(* IEC 61131-3 sources: plc-process-lib/tools/demo/src/POUs/FB_DemoLevelLoop, 2 files *)

(* ---- FB_DemoLevelLoop.decl.st ---- *)
// Назначение: сценарий A демонстрационного прогона — контур уровня по примеру 17.3 контракта:
//             LT (PL.FB_AnalogInput, 4–20 мА, 0..5 м) -> LIC (PL.FB_PID, Direct, обратный расчёт
//             по фактическому заданию ПЧ) -> насос с ПЧ (PL.FB_MotorVfd, мин. 20 %). Объект —
//             модель ёмкости на ST: баланс объёма, подача насоса пропорциональна скорости, ПЧ
//             разгоняется с рампой. Сценарий: 5 с — пуск насоса (слежение ПИД снимается без
//             рывка); 40 с — задание 2,5 -> 1,5 м (выход упирается в 100 %, интегратор не
//             накапливается); 95 с — приток 120 -> 210 м3/ч. Ёмкость и параметры вымышленные.
//             Коды событий: 1 — пуск насоса, 2 — ступень задания, 3 — ступень притока.
// Автор:      kr0nsch
// Версия:     0.1.0
// Документ:   docs/API.md, пример 17.3; tools/demo/README.md
FUNCTION_BLOCK FB_DemoLevelLoop
VAR_INPUT
    lrT_s  : LREAL;   // время от старта сценария, с
    lrDt_s : LREAL;   // шаг времени этого цикла, с
END_VAR
VAR_OUTPUT
    xDone : BOOL;     // сценарий завершён, журнал записан
END_VAR
VAR CONSTANT
    LEVEL_SPAN_M   : REAL := 5.0;       // шкала датчика: 4 мА = 0 м, 20 мА = 5 м
    MA_LO          : REAL := 4.0;       // ток начала шкалы, мА
    MA_SPAN        : REAL := 16.0;      // диапазон тока шкалы, мА
    AREA_M2        : LREAL := 1.5;      // площадь сечения ёмкости, м2
    LEVEL0_M       : LREAL := 2.3;      // начальный уровень, м
    Q_PUMP_MAX_M3H : REAL := 300.0;     // подача насоса при 100 % скорости, м3/ч (линейная модель)
    Q_IN_BASE_M3H  : REAL := 120.0;     // приток до возмущения, м3/ч
    Q_IN_SURGE_M3H : REAL := 210.0;     // приток после возмущения, м3/ч
    VFD_RAMP_PCTPS : REAL := 25.0;      // рампа ПЧ (модель привода), %/с
    S_PER_H        : LREAL := 3600.0;   // секунд в часе
    PCT_FULL       : REAL := 100.0;     // 100 %
    SP0_M          : REAL := 2.5;       // задание до ступени, м
    SP1_M          : REAL := 1.5;       // задание после ступени, м
    T_START_S      : LREAL := 5.0;      // пуск насоса (xAutoRun), с
    T_SP_STEP_S    : LREAL := 40.0;     // ступень задания, с
    T_SURGE_S      : LREAL := 95.0;     // ступень притока, с
    PID_KP         : REAL := 12.0;      // коэффициент усиления, %/%
    PID_TI_S       : REAL := 80.0;      // время интегрирования, с
    SPEED_MIN_PCT  : REAL := 20.0;      // мин. задание ПЧ в работе, %
    SCENARIO       : INT := 1;          // номер сценария в журнале событий
    EV_START       : INT := 1;          // событие: пуск насоса
    EV_SP_STEP     : INT := 2;          // событие: ступень задания
    EV_SURGE       : INT := 3;          // событие: ступень притока
END_VAR
VAR
    // устройства библиотеки, обмен — через структуры команд, Cfg и Retain, как в приложении
    fbLt          : PL.FB_AnalogInput;    // LT: датчик уровня
    stLtCmd       : PL.ST_AnalogInputCmd; // его команды
    stLtCfg       : PL.ST_AnalogInputCfg; // его Cfg
    fbLic         : PL.FB_PID;            // LIC: регулятор уровня
    stLicCmd      : PL.ST_PidCmd;         // его команды (задание оператора)
    stLicRet      : PL.ST_DeviceRetain;   // его режим
    stLicCfg      : PL.ST_PidCfg;         // его Cfg
    fbPump        : PL.FB_MotorVfd;       // насос с ПЧ
    stPumpCmd     : PL.ST_MotorCmd;       // его команды
    stPumpRet     : PL.ST_DeviceRetain;   // его режим и счётчики
    stPumpCfg     : PL.ST_MotorCfg;       // его Cfg
    // модель объекта
    lrLevel_m     : LREAL;                // уровень в ёмкости, м
    rSpeedAct_pct : REAL;                 // скорость ПЧ, %
    rQin_m3h      : REAL;                 // приток, м3/ч
    rQout_m3h     : REAL;                 // отбор насосом, м3/ч
    rLevel_mA     : REAL;                 // ток датчика уровня, мА
    // контур
    xLeadAuto     : BOOL;                 // насос в Auto и работает (прошлый цикл): ПИД не следит
    rLeadRef_pct  : REAL;                 // задание ПЧ прошлого цикла, %
    // сценарий и журнал
    xInit         : BOOL;                 // Cfg и начальное состояние заданы
    xStartDone    : BOOL;                 // пуск насоса выполнен
    xSpDone       : BOOL;                 // ступень задания выполнена
    xSurgeDone    : BOOL;                 // ступень притока выполнена
    lrNextLog_s   : LREAL;                // время следующей записи журнала, с
    uiIdx         : UINT;                 // индекс записи журнала
END_VAR

(* ---- FB_DemoLevelLoop.impl.st ---- *)
IF NOT xInit THEN
    xInit := TRUE;
    stLtCfg.rRangeHi_eu := LEVEL_SPAN_M;
    stLicCfg.eAction := PL.E_PidAction.Direct;          // уровень выше задания -> насос быстрее
    stLicCfg.rKp := PID_KP;
    stLicCfg.rTi_s := PID_TI_S;
    stLicCfg.rPvMax_eu := LEVEL_SPAN_M;
    stLicCfg.rSpMax_eu := LEVEL_SPAN_M;
    stLicCfg.xUseOutAct := TRUE;                        // обратный расчёт по фактическому заданию ПЧ
    stLicRet.eRemoteMode := PL.E_DeviceMode.Auto;
    stLicCmd.rSp_eu := SP0_M;
    stPumpCfg.stVfd.rSpeedMin_pct := SPEED_MIN_PCT;
    stPumpRet.eRemoteMode := PL.E_DeviceMode.Auto;
    lrLevel_m := LEVEL0_M;
END_IF
IF xDone THEN
    RETURN;
END_IF

// Сценарий: пуск насоса, ступень задания, ступень притока
IF lrT_s >= T_START_S AND NOT xStartDone THEN
    xStartDone := TRUE;
    fbPump.xAutoRun := TRUE;
    F_DemoEvent(lrT_s := lrT_s, iScenario := SCENARIO, iCode := EV_START);
END_IF
IF lrT_s >= T_SP_STEP_S AND NOT xSpDone THEN
    xSpDone := TRUE;
    stLicCmd.rSp_eu := SP1_M;
    F_DemoEvent(lrT_s := lrT_s, iScenario := SCENARIO, iCode := EV_SP_STEP);
END_IF
IF lrT_s >= T_SURGE_S AND NOT xSurgeDone THEN
    xSurgeDone := TRUE;
    F_DemoEvent(lrT_s := lrT_s, iScenario := SCENARIO, iCode := EV_SURGE);
END_IF
rQin_m3h := SEL(xSurgeDone, Q_IN_BASE_M3H, Q_IN_SURGE_M3H);

// Датчик уровня: уровень модели -> ток 4–20 мА
rLevel_mA := MA_LO + MA_SPAN * LREAL_TO_REAL(lrLevel_m) / LEVEL_SPAN_M;

// Контур по примеру 17.3 контракта: насос (прошлый вызов) -> AI -> ПИД -> задание ПЧ -> ПЧ.
// Пока насос не в Auto-работе, ПИД следит за заданием ПЧ: пуск и переходы режимов без рывка
xLeadAuto := fbPump.SpeedAutoActive;
rLeadRef_pct := fbPump.SpeedRef;
fbLt(rIn := rLevel_mA, stCmd := stLtCmd, stCfg := stLtCfg);
fbLic(rPv_eu := fbLt.rValue_eu, xPvValid := fbLt.xValid, xTrack := NOT xLeadAuto, rTrack_pct := rLeadRef_pct,
      rOutAct_pct := rLeadRef_pct, stCmd := stLicCmd, stRetain := stLicRet, stCfg := stLicCfg);
fbPump.rSpeedSpAuto_pct := fbLic.rOut_pct;
fbPump(stCmd := stPumpCmd, stRetain := stPumpRet, stCfg := stPumpCfg);

// Модель ПЧ: работает по команде, скорость идёт к заданию с рампой привода
rSpeedAct_pct := PL.F_RateLimit(rCurrent := rSpeedAct_pct,
                                rTarget := SEL(fbPump.xQRun, 0.0, fbPump.rSpeedRef_pct),
                                rRateUp_ups := VFD_RAMP_PCTPS, rRateDown_ups := VFD_RAMP_PCTPS,
                                lrDt_s := lrDt_s);
fbPump.xVfdRunning := fbPump.xQRun;
fbPump.rSpeedAct_pct := rSpeedAct_pct;

// Модель ёмкости: баланс объёма
rQout_m3h := Q_PUMP_MAX_M3H * rSpeedAct_pct / PCT_FULL;
lrLevel_m := lrLevel_m + REAL_TO_LREAL(rQin_m3h - rQout_m3h) / S_PER_H / AREA_M2 * lrDt_s;
lrLevel_m := LIMIT(0.0, lrLevel_m, REAL_TO_LREAL(LEVEL_SPAN_M));

// Журнал с периодом LOOP_LOG_PERIOD_S
IF lrT_s >= lrNextLog_s AND GVL_DemoLog.uiLoopN < GVL_DemoConst.LOOP_LOG_N THEN
    uiIdx := GVL_DemoLog.uiLoopN;
    GVL_DemoLog.arLoopT_s[uiIdx] := LREAL_TO_REAL(lrT_s);
    GVL_DemoLog.arLoopLevel_m[uiIdx] := LREAL_TO_REAL(lrLevel_m);
    GVL_DemoLog.arLoopPv_m[uiIdx] := fbLt.rValue_eu;
    GVL_DemoLog.arLoopSp_m[uiIdx] := fbLic.stSts.rSp_eu;
    GVL_DemoLog.arLoopOut_pct[uiIdx] := fbLic.rOut_pct;
    GVL_DemoLog.arLoopP_pct[uiIdx] := fbLic.stSts.rP_pct;
    GVL_DemoLog.arLoopI_pct[uiIdx] := fbLic.stSts.rI_pct;
    GVL_DemoLog.arLoopRef_pct[uiIdx] := fbPump.rSpeedRef_pct;
    GVL_DemoLog.arLoopAct_pct[uiIdx] := rSpeedAct_pct;
    GVL_DemoLog.arLoopQin_m3h[uiIdx] := rQin_m3h;
    GVL_DemoLog.arLoopQout_m3h[uiIdx] := rQout_m3h;
    GVL_DemoLog.aiLoopMotor[uiIdx] := TO_INT(fbPump.stSts.eState);
    GVL_DemoLog.awLoopPidSts[uiIdx] := fbLic.stSts.stCommon.wStatus;
    GVL_DemoLog.uiLoopN := uiIdx + 1;
    lrNextLog_s := lrNextLog_s + GVL_DemoConst.LOOP_LOG_PERIOD_S;
END_IF
xDone := lrT_s >= GVL_DemoConst.LOOP_DURATION_S;
